(* IEC 61131-3 sources: llm-plc-st-eval/data/definitivo/gemini-3.1-pro-preview/B5/zero_shot, 3 files *)

(* ---- ejec_1.st ---- *)
```iecst
FUNCTION_BLOCK FB_Ventilador
VAR_INPUT
    quemadorOn : BOOL; // Indica si el quemador está encendido
END_VAR
VAR_OUTPUT
    ventilador : BOOL; // Controla el estado del ventilador
END_VAR
VAR
    temporizadorTOF : TOF; // Temporizador de retardo a la desconexión (Off-Delay)
END_VAR

// El temporizador TOF mantiene su salida Q en TRUE mientras IN sea TRUE,
// y la mantiene 30 segundos adicionales después de que IN pase a FALSE.
temporizadorTOF(IN := quemadorOn, PT := T#30S);

// Asignación directa de la salida del temporizador al ventilador
ventilador := temporizadorTOF.Q;

END_FUNCTION_BLOCK
```

(* ---- ejec_2.st ---- *)
```iecst
FUNCTION_BLOCK FB_Ventilador
VAR_INPUT
    quemadorOn : BOOL; // Indica si el quemador está encendido
END_VAR

VAR_OUTPUT
    ventilador : BOOL; // Comando de encendido para el ventilador
END_VAR

VAR
    temporizadorTOF : TOF; // Temporizador de retardo a la desconexión (Off-Delay)
END_VAR

// Configuración y ejecución del temporizador
// Si quemadorOn es TRUE, la salida Q es TRUE inmediatamente.
// Cuando quemadorOn pasa a FALSE, Q se mantiene TRUE durante el tiempo PT (30s) y luego pasa a FALSE.
temporizadorTOF(IN := quemadorOn, PT := T#30S);

// Asignación del estado del temporizador a la salida del ventilador
ventilador := temporizadorTOF.Q;

END_FUNCTION_BLOCK
```

(* ---- ejec_3.st ---- *)
```iecst
FUNCTION_BLOCK FB_Ventilador
VAR_INPUT
    quemadorOn : BOOL; // Indica si el quemador está encendido
END_VAR
VAR_OUTPUT
    ventilador : BOOL; // Controla el estado del ventilador
END_VAR
VAR
    timerTOF : TOF; // Temporizador de retardo a la desconexión (Off-Delay)
END_VAR

// Llamada al temporizador:
// Mientras IN es TRUE, Q es TRUE.
// Cuando IN pasa a FALSE, Q se mantiene TRUE durante el tiempo PT (30s) y luego pasa a FALSE.
timerTOF(IN := quemadorOn, PT := T#30S);

// Asignación de la salida del temporizador al ventilador
ventilador := timerTOF.Q;

END_FUNCTION_BLOCK
```
